// TIA Portal V20 export
// export: Created 2026-10-20T12:46:08.391772Z, ExportSetting WithDefaults, DisplayName Totally Integrated Automation Portal, DisplayVersion V20 Update 6, DisplayName TIA Portal Openness, DisplayVersion V20 Update 6, DisplayName TIA Portal Version Control Interface, DisplayVersion V20 Update 6, DisplayName SINAMICS Startdrive Advanced, DisplayVersion V20 SP1, DisplayName SINAMICS Startdrive G130, G150, S120, S150, SINAMICS MV, G220, S200, S210, DisplayVersion V20 SP1, DisplayName SINAMICS Startdrive G110M, G120, G120C, G120D, G120P, G115D, DisplayVersion V20 SP1, DisplayName STEP 7 Professional, DisplayVersion V20 Update 6, DisplayName STEP 7 Safety, DisplayVersion V20 Update 2, DisplayName WinCC Basic/Comfort/Advanced, DisplayVersion V20 Update 6, DisplayName WinCC Unified, DisplayVersion V20 Update 6
DATA_BLOCK "PopUps_DB_1"   // DB20
{ S7_Optimized_Access := 'TRUE' }
VERSION : 0.1
// stored: AutoNumber true, DBAccessibleFromOPCUA true, IsOnlyStoredInLoadMemory false, IsRetainMemResEnabled false, IsWriteProtectedInAS false, MemoryReserve 100
   VAR
      Buffer_Cnv_Settings_1 : Array[1..5] of "Buffer_Cnv_Settings";
      Buffer_Cnv_Settings_2 { S7_SetPoint := 'True'} : Array[1..5] of "Buffer_Cnv_Settings";
      ECnv_Settings { S7_SetPoint := 'True'} : Array[1..5] of "ECnv_Settings";
      VTD_Settings { S7_SetPoint := 'True'} : Array[1..5] of "VTD_Settings";
      Shuttle_MQTT_Settings { S7_SetPoint := 'True'} : "MQTT_Settings";
      Sick_Lector_Reseult : Array[1..5] of String;
      Save_Settings { S7_SetPoint := 'True'} : Array[1..5] of Bool;
      Absolute_Encoder : Array[1..5] of Struct
         AE_Control_Word_1 : UInt;
         AE_Control_Word_2 : UInt;
         AE_Status_1 : UInt;
         AE_Status_2 : UInt;
         AE_Position_1 : DInt;
         AE_Position_2 : DInt;
         AE_Speed : Int;
      END_STRUCT;
      Lector_Barcode : Array[1..5] of Struct
         BCD_Test_Comm : Bool;
         BCD_Disable_Trigger : Bool;
         BCD_Enable_Trigger : Bool;
         BCD_Execute_Function : Bool;
         BCD_Test_Ok : Bool;
         BCD_Error : Bool;
         BCD_RdDone : Bool;
         BCD_ReqDone : Bool;
         BCD_ReqBusy : Bool;
         Lector_Reseult : String;
      END_STRUCT;
      Linear_Encoder : Array[1..5] of Struct
         LE_X_Unsafe_Position : DInt;
         LE_Speed : Int;
         LE_Warnings : Int;
         LE_Bypass : Bool;
         LE_Status : UInt;
      END_STRUCT;
      Trend : Array[1..5] of Struct
         Motor_SetPoint : UInt;
         Motor_Actual_Current : Real;
         Motor_Actual_Speed : UInt;
      END_STRUCT;
   END_VAR
BEGIN
   Shuttle_MQTT_Settings.MQTT_Con_Params.hwId := 64;
   Shuttle_MQTT_Settings.MQTT_Con_Params.broker := '10.0.34.2';
   Shuttle_MQTT_Settings.Client_ID := WSTRING#'PLC';
   Shuttle_MQTT_Settings.Username := WSTRING#'Devin';
   Shuttle_MQTT_Settings.Password := WSTRING#'1';
   Shuttle_MQTT_Settings.Retain := TRUE;
END_DATA_BLOCK
